Staubli VAL3: HMI_cycle.dtx

mdesc mNomSpeed
bool bReset
bool bStart
bool bHold
bool bEnd
bool bStop
bool bBack
bool bToHome
bool bClearErr
string sState
string sCapacity
string sAvgCapacity
string sBestCapacity
string sProgCode
num nLastProg
string sTrajStatus
string sLib
num nLastLib
bool bRotBack
